Fanuc KAREL source: KD00061.KL

PROGRAM KD00061
%NOLOCKGROUP
VAR
  I: INTEGER
  J: INTEGER
  B: BOOLEAN
  R: REAL
  S: STRING[80]
BEGIN
  CONDITION[1]:
  WHEN DIN[1] = ON DO
    DISABLE CONDITION[1]
  ENDCONDITION
END KD00061
